(* IEC 61131-3 sources: AgenticPLC_Editor/AgenticPLC-editor/resources/strucpp/libs/sources/additional-function-blocks, 6 files *)

(* ---- derivative.st ---- *)
(* Additional Function Blocks: DERIVATIVE                                *)
(* Source carried verbatim from MatIEC's lib/derivative_st.txt.          *)
(* Original header preserved for traceability:                           *)
(*   "Following taken directly from the IEC 61131.3 draft standard"      *)
(*   "FINAL DRAFT - IEC 61131-3, 2nd Ed. (2001-12-10)"                   *)

FUNCTION_BLOCK DERIVATIVE
  VAR_INPUT
    RUN   : BOOL ;          (* 0 = reset                  *)
    XIN   : REAL ;          (* Input to be differentiated *)
    CYCLE : TIME ;          (* Sampling period            *)
  END_VAR
  VAR_OUTPUT
    XOUT : REAL ;           (* Differentiated output      *)
  END_VAR
  VAR
    X1 : REAL ;
    X2 : REAL ;
    X3 : REAL ;
  END_VAR

  IF RUN THEN
    XOUT := (3.0 * (XIN - X3) + X1 - X2) / (10.0 * TIME_TO_REAL(CYCLE)) ;
    X3 := X2 ;
    X2 := X1 ;
    X1 := XIN ;
  ELSE
    XOUT := 0.0 ;
    X1 := XIN ;
    X2 := XIN ;
    X3 := XIN ;
  END_IF ;
END_FUNCTION_BLOCK

(* ---- hysteresis.st ---- *)
(* Additional Function Blocks: HYSTERESIS                                *)
(* Source carried verbatim from MatIEC's lib/hysteresis_st.txt.          *)
(* Original header preserved for traceability:                           *)
(*   "Following taken directly from the IEC 61131.3 draft standard"      *)
(*   "FINAL DRAFT - IEC 61131-3, 2nd Ed. (2001-12-10)"                   *)
(*                                                                        *)
(* Boolean hysteresis on the difference of two REAL inputs (XIN1 - XIN2). *)

FUNCTION_BLOCK HYSTERESIS
  VAR_INPUT
    XIN1 : REAL ;
    XIN2 : REAL ;
    EPS  : REAL ;
  END_VAR
  VAR_OUTPUT
    Q : BOOL := FALSE ;
  END_VAR

  IF Q THEN
    IF XIN1 < (XIN2 - EPS) THEN
      Q := FALSE ;
    END_IF ;
  ELSIF XIN1 > (XIN2 + EPS) THEN
    Q := TRUE ;
  END_IF ;
END_FUNCTION_BLOCK

(* ---- integral.st ---- *)
(* Additional Function Blocks: INTEGRAL                                  *)
(* Source carried verbatim from MatIEC's lib/integral_st.txt.            *)
(* Original header preserved for traceability:                           *)
(*   "Following taken directly from the IEC 61131.3 draft standard"      *)
(*   "FINAL DRAFT - IEC 61131-3, 2nd Ed. (2001-12-10)"                   *)

FUNCTION_BLOCK INTEGRAL
  VAR_INPUT
    RUN   : BOOL ;       (* 1 = integrate, 0 = hold *)
    R1    : BOOL ;       (* Overriding reset        *)
    XIN   : REAL ;       (* Input variable          *)
    X0    : REAL ;       (* Initial value           *)
    CYCLE : TIME ;       (* Sampling period         *)
  END_VAR
  VAR_OUTPUT
    Q    : BOOL ;        (* NOT R1                  *)
    XOUT : REAL ;        (* Integrated output       *)
  END_VAR

  Q := NOT R1 ;
  IF R1 THEN
    XOUT := X0 ;
  ELSIF RUN THEN
    XOUT := XOUT + XIN * TIME_TO_REAL(CYCLE) ;
  END_IF ;
END_FUNCTION_BLOCK

(* ---- pid.st ---- *)
(* Additional Function Blocks: PID                                       *)
(* Source carried verbatim from MatIEC's lib/pid_st.txt.                 *)
(* Original header preserved for traceability:                           *)
(*   "Following taken directly from the IEC 61131.3 draft standard"      *)
(*   "FINAL DRAFT - IEC 61131-3, 2nd Ed. (2001-12-10)"                   *)
(*                                                                        *)
(* Depends on INTEGRAL and DERIVATIVE FBs declared elsewhere in this lib. *)

FUNCTION_BLOCK PID
  VAR_INPUT
    AUTO  : BOOL ;       (* 0 - manual , 1 - automatic *)
    PV    : REAL ;       (* Process variable *)
    SP    : REAL ;       (* Set point *)
    X0    : REAL ;       (* Manual output adjustment - typically from transfer station *)
    KP    : REAL ;       (* Proportionality constant *)
    TR    : REAL ;       (* Reset time *)
    TD    : REAL ;       (* Derivative time constant *)
    CYCLE : TIME ;       (* Sampling period *)
  END_VAR
  VAR_OUTPUT
    XOUT : REAL ;
  END_VAR
  VAR
    ERROR : REAL ;        (* PV - SP *)
    ITERM : INTEGRAL ;    (* FB for integral term  *)
    DTERM : DERIVATIVE ;  (* FB for derivative term *)
  END_VAR

  ERROR := PV - SP ;
  (*** Adjust ITERM so that XOUT := X0 when AUTO = 0 ***)
  ITERM (RUN := AUTO, R1 := NOT AUTO, XIN := ERROR,
         X0 := TR * (X0 - ERROR), CYCLE := CYCLE) ;
  DTERM (RUN := AUTO, XIN := ERROR, CYCLE := CYCLE) ;
  XOUT := KP * (ERROR + ITERM.XOUT / TR + DTERM.XOUT * TD) ;
END_FUNCTION_BLOCK

(* ---- ramp.st ---- *)
(* Additional Function Blocks: RAMP                                      *)
(* Source carried verbatim from MatIEC's lib/ramp_st.txt.                *)
(* Original header preserved for traceability:                           *)
(*   "Following taken directly from the IEC 61131.3 draft standard"      *)
(*   "FINAL DRAFT - IEC 61131-3, 2nd Ed. (2001-12-10)"                   *)

FUNCTION_BLOCK RAMP
  VAR_INPUT
    RUN   : BOOL ;       (* 0 - track X0, 1 - ramp to/track X1 *)
    X0    : REAL ;
    X1    : REAL ;
    TR    : TIME ;       (* Ramp duration *)
    CYCLE : TIME ;       (* Sampling period *)
  END_VAR
  VAR_OUTPUT
    BUSY : BOOL ;        (* BUSY = 1 during ramping period *)
    XOUT : REAL := 0.0 ;
  END_VAR
  VAR
    XI : REAL ;          (* Initial value *)
    T  : TIME := T#0s ;  (* Elapsed time of ramp *)
  END_VAR

  BUSY := RUN ;
  IF RUN THEN
    IF T >= TR THEN
      BUSY := FALSE ;
      XOUT := X1 ;
    ELSE
      XOUT := XI + (X1 - XI) * TIME_TO_REAL(T) / TIME_TO_REAL(TR) ;
      T := T + CYCLE ;
    END_IF ;
  ELSE
    XOUT := X0 ;
    XI := X0 ;
    T := T#0s ;
  END_IF ;
END_FUNCTION_BLOCK

(* ---- rtc.st ---- *)
(* Additional Function Blocks: RTC                                       *)
(* Source ported verbatim from MatIEC's lib/rtc.txt with one substitution: *)
(* the MatIEC pragma `{__SET_VAR(data__->,CURRENT_TIME,,__CURRENT_TIME)}`  *)
(* read MatIEC's `__CURRENT_TIME` global, which serves the same purpose as *)
(* STruC++'s TIME() — monotonic scan-cycle time, hardware agnostic. We     *)
(* substitute TO_DT(TIME()) so the same int64 tick value lands in a DT-    *)
(* typed local. STruC++ requires an explicit conversion where MatIEC's     *)
(* pragma did a raw bit-copy; behaviour is otherwise identical.            *)
(*                                                                        *)
(* Original MatIEC documentation:                                          *)
(*                                                                        *)
(*   RTC - Real-time clock                                                *)
(*                                                                        *)
(*   Q is a copy of IN.                                                    *)
(*                                                                        *)
(*   When IN = FALSE, CDT is the current "tick" time exposed by the       *)
(*   runtime as a DT.                                                      *)
(*                                                                        *)
(*   When IN changes from FALSE to TRUE, PDT is stored. As long as IN is   *)
(*   TRUE, CDT is equal to PDT + the amount of time since PDT was loaded. *)

FUNCTION_BLOCK RTC
  VAR_INPUT
    IN  : BOOL ;                  (* 0 - current time, 1 - load time from PDT *)
    PDT : DT ;                    (* Preset datetime *)
  END_VAR
  VAR_OUTPUT
    Q   : BOOL := FALSE ;         (* Copy of IN *)
    CDT : DT ;                    (* Datetime, current or relative to PDT *)
  END_VAR

  VAR
    PREV_IN      : BOOL := FALSE ;
    OFFSET       : TIME ;
    CURRENT_TIME : DT ;
  END_VAR

  CURRENT_TIME := TO_DT(TIME()) ;

  IF IN THEN
    IF NOT PREV_IN THEN
      OFFSET := PDT - CURRENT_TIME ;
    END_IF ;

    (* PDT + time since PDT was loaded *)
    CDT := CURRENT_TIME + OFFSET ;
  ELSE
    CDT := CURRENT_TIME ;
  END_IF ;

  Q := IN ;
  PREV_IN := IN ;
END_FUNCTION_BLOCK
